(* IEC 61131-3 sources: RVM_Dijital_Ikiz_ModelveOtomasyon_BitirmeProjesi/simulasyon_unity/plc, 14 files *)

(* ---- ST_RVMInput106.st ---- *)
TYPE ST_RVMInput106 :
STRUCT
    uiUnityProtokol : UINT := 106;
    udiUnityOturumu : UDINT := 0;
    udiUnitySayaci : UDINT := 0;
    udiKomutKimligi : UDINT := 0;
    uiOperatorKomutu : UINT := 0;
    xGiris : BOOL := FALSE;
    xTanima : BOOL := FALSE;
    xKiriciGiris : BOOL := FALSE;
    xKirildi : BOOL := FALSE;
    xHazneDolu : BOOL := FALSE;
    xBosaltildi : BOOL := FALSE;
    xKapakAcik : BOOL := FALSE;
    xKapakKapali : BOOL := FALSE;
    xYolBos : BOOL := FALSE;
    xMetalAlgilandi : BOOL := FALSE;
    xSikisma : BOOL := FALSE;
    xAcilStop : BOOL := FALSE;
    xKutuPetDolu : BOOL := FALSE;
    xKutuAluminyumDolu : BOOL := FALSE;
    xKutuCamDolu : BOOL := FALSE;
    rKutleGram : REAL := 0.0;
    rOptikGecirgenlik : REAL := 0.0;
    rBoyMetre : REAL := 0.0;
    rHazneKonumu : REAL := 0.0;
    rGercekBantHizi : REAL := 0.0;
    rGercekKiriciDevri : REAL := 0.0;
    uiBosaltilanKutu : UINT := 0;
    udiUrunKimligi : UDINT := 0;
    uiOperatorParametresi : UINT := 0;
    udiGorulenPlcOturumu : UDINT := 0;
    udiNesneOnayi : UDINT := 0;
    uiNesneSonucu : UINT := 0;
    udiNesneUrunKimligi : UDINT := 0;
    uiPlantVeriKaynagi : UINT := 0;
    xPlantVerisiGecerli : BOOL := FALSE;
    udiGoruntuOnayi : UDINT := 0;
    udiGoruntuUrunu : UDINT := 0;
    udiGoruntuPlcOturumu : UDINT := 0;
    udiGoruntuUnityOturumu : UDINT := 0;
    xGoruntuGecerli : BOOL := FALSE;
    xGoruntuNesneVar : BOOL := FALSE;
    rGoruntuBoy : REAL := 0;
    rGoruntuEn : REAL := 0;
    rGoruntuDoluluk : REAL := 0;
    rGoruntuYasiMs : REAL := 0;
    xOlcumTartiGecerli : BOOL;
    xOlcumProbGecerli : BOOL;
    rOlcumYansima : REAL;
    rOlcumMetal : REAL;
    rOlcumManyetik : REAL;
END_STRUCT
END_TYPE

(* ---- ST_RVMOperator106.st ---- *)
TYPE ST_RVMOperator106 :
STRUCT
    xBaslat : BOOL := FALSE;
    xDurdur : BOOL := FALSE;
    xSifirla : BOOL := FALSE;
    xNesneEkle : BOOL := FALSE;
    xModUygula : BOOL := FALSE;
    xAcilStop : BOOL := FALSE;
    uiSeciliNesne : UINT := 1;
    uiSeciliMod : UINT := 1;
END_STRUCT
END_TYPE

(* ---- ST_RVMOutput106.st ---- *)
TYPE ST_RVMOutput106 :
STRUCT
    uiProtokolSurumu : UINT := 106;
    udiPlcSayaci : UDINT := 0;
    udiUnityOnayOturumu : UDINT := 0;
    udiGirisOnayi : UDINT := 0;
    udiKomutOnayi : UDINT := 0;
    udiIslemKimligi : UDINT := 0;
    uiDurum : UINT := 0;
    uiHataKodu : UINT := 0;
    uiTaninmisMalzeme : UINT := 0;
    uiHedefKutu : UINT := 0;
    xCalismaIzni : BOOL := FALSE;
    xKonveyorIleri : BOOL := FALSE;
    xKonveyorGeri : BOOL := FALSE;
    xKiriciCalis : BOOL := FALSE;
    xHazneHareket : BOOL := FALSE;
    xKapakAc : BOOL := FALSE;
    xTanimaOnayi : BOOL := FALSE;
    rBantHizi : REAL := 0.85;
    rKiriciDevri : REAL := 120.0;
    rHazneHizi : REAL := 1.5;
    rHazneHedefi : REAL := 0.0;
    rKapakAcisi : REAL := 75.0;
    udiPetSayaci : UDINT := 0;
    udiAluminyumSayaci : UDINT := 0;
    udiCamSayaci : UDINT := 0;
    udiReddedilenSayaci : UDINT := 0;
    udiPlcOturumu : UDINT := 0;
    uiKomutDurumu : UINT := 0;
    uiKomutNedeni : UINT := 0;
    udiPlcOperatorKomutKimligi : UDINT := 0;
    uiPlcOperatorKomutu : UINT := 0;
    uiPlcKomutDurumu : UINT := 0;
    uiPlcKomutNedeni : UINT := 0;
    uiSonKomutKaynagi : UINT := 0;
    udiNesneIstegi : UDINT := 0;
    uiNesneProfili : UINT := 0;
    xNesneIstegiEtkin : BOOL := FALSE;
    uiVeriModu : UINT := 1;
    uiDesteklenenModlar : UINT := 2;
    udiCikisBaslangic : UDINT := 0;
    udiCikisBitis : UDINT := 0;
    udiGoruntuIstegi : UDINT := 0;
    uiGoruntuKarari : UINT := 0;
END_STRUCT
END_TYPE

(* ---- GVL_RVMKalici.st ---- *)
{attribute 'qualified_only'}
VAR_GLOBAL PERSISTENT RETAIN
    udiOturum : UDINT;
END_VAR

(* ---- GVL_RVMOperator.st ---- *)
{attribute 'qualified_only'}
VAR_GLOBAL
    xBaslat : BOOL := FALSE;
    xDurdur : BOOL := FALSE;
    xSifirla : BOOL := FALSE;
    xNesneEkle : BOOL := FALSE;
    xModUygula : BOOL := FALSE;
    xAcilStop : BOOL := FALSE;
    uiSeciliNesne : UINT := 1;
    uiSeciliMod : UINT := 1;
END_VAR

(* ---- GVL_RVMUnity.st ---- *)
{attribute 'qualified_only'}
VAR_GLOBAL
    {attribute 'symbol' := 'readwrite'}
    uiUnityProtokol : UINT := 106;
    {attribute 'symbol' := 'readwrite'}
    udiUnityOturumu : UDINT := 0;
    {attribute 'symbol' := 'readwrite'}
    udiUnitySayaci : UDINT := 0;
    {attribute 'symbol' := 'readwrite'}
    udiKomutKimligi : UDINT := 0;
    {attribute 'symbol' := 'readwrite'}
    uiOperatorKomutu : UINT := 0;
    {attribute 'symbol' := 'readwrite'}
    xGiris : BOOL := FALSE;
    {attribute 'symbol' := 'readwrite'}
    xTanima : BOOL := FALSE;
    {attribute 'symbol' := 'readwrite'}
    xKiriciGiris : BOOL := FALSE;
    {attribute 'symbol' := 'readwrite'}
    xKirildi : BOOL := FALSE;
    {attribute 'symbol' := 'readwrite'}
    xHazneDolu : BOOL := FALSE;
    {attribute 'symbol' := 'readwrite'}
    xBosaltildi : BOOL := FALSE;
    {attribute 'symbol' := 'readwrite'}
    xKapakAcik : BOOL := FALSE;
    {attribute 'symbol' := 'readwrite'}
    xKapakKapali : BOOL := FALSE;
    {attribute 'symbol' := 'readwrite'}
    xYolBos : BOOL := FALSE;
    {attribute 'symbol' := 'readwrite'}
    xMetalAlgilandi : BOOL := FALSE;
    {attribute 'symbol' := 'readwrite'}
    xSikisma : BOOL := FALSE;
    {attribute 'symbol' := 'readwrite'}
    xAcilStop : BOOL := FALSE;
    {attribute 'symbol' := 'readwrite'}
    xKutuPetDolu : BOOL := FALSE;
    {attribute 'symbol' := 'readwrite'}
    xKutuAluminyumDolu : BOOL := FALSE;
    {attribute 'symbol' := 'readwrite'}
    xKutuCamDolu : BOOL := FALSE;
    {attribute 'symbol' := 'readwrite'}
    rKutleGram : REAL := 0.0;
    {attribute 'symbol' := 'readwrite'}
    rOptikGecirgenlik : REAL := 0.0;
    {attribute 'symbol' := 'readwrite'}
    rBoyMetre : REAL := 0.0;
    {attribute 'symbol' := 'readwrite'}
    rHazneKonumu : REAL := 0.0;
    {attribute 'symbol' := 'readwrite'}
    rGercekBantHizi : REAL := 0.0;
    {attribute 'symbol' := 'readwrite'}
    rGercekKiriciDevri : REAL := 0.0;
    {attribute 'symbol' := 'readwrite'}
    uiBosaltilanKutu : UINT := 0;
    {attribute 'symbol' := 'readwrite'}
    udiUrunKimligi : UDINT := 0;
    {attribute 'symbol' := 'read'}
    uiProtokolSurumu : UINT := 106;
    {attribute 'symbol' := 'read'}
    udiPlcSayaci : UDINT := 0;
    {attribute 'symbol' := 'read'}
    udiUnityOnayOturumu : UDINT := 0;
    {attribute 'symbol' := 'read'}
    udiGirisOnayi : UDINT := 0;
    {attribute 'symbol' := 'read'}
    udiKomutOnayi : UDINT := 0;
    {attribute 'symbol' := 'read'}
    udiIslemKimligi : UDINT := 0;
    {attribute 'symbol' := 'read'}
    uiDurum : UINT := 0;
    {attribute 'symbol' := 'read'}
    uiHataKodu : UINT := 0;
    {attribute 'symbol' := 'read'}
    uiTaninmisMalzeme : UINT := 0;
    {attribute 'symbol' := 'read'}
    uiHedefKutu : UINT := 0;
    {attribute 'symbol' := 'read'}
    xCalismaIzni : BOOL := FALSE;
    {attribute 'symbol' := 'read'}
    xKonveyorIleri : BOOL := FALSE;
    {attribute 'symbol' := 'read'}
    xKonveyorGeri : BOOL := FALSE;
    {attribute 'symbol' := 'read'}
    xKiriciCalis : BOOL := FALSE;
    {attribute 'symbol' := 'read'}
    xHazneHareket : BOOL := FALSE;
    {attribute 'symbol' := 'read'}
    xKapakAc : BOOL := FALSE;
    {attribute 'symbol' := 'read'}
    xTanimaOnayi : BOOL := FALSE;
    {attribute 'symbol' := 'read'}
    rBantHizi : REAL := 0.85;
    {attribute 'symbol' := 'read'}
    rKiriciDevri : REAL := 120.0;
    {attribute 'symbol' := 'read'}
    rHazneHizi : REAL := 1.5;
    {attribute 'symbol' := 'read'}
    rHazneHedefi : REAL := 0.0;
    {attribute 'symbol' := 'read'}
    rKapakAcisi : REAL := 75.0;
    {attribute 'symbol' := 'read'}
    udiPetSayaci : UDINT := 0;
    {attribute 'symbol' := 'read'}
    udiAluminyumSayaci : UDINT := 0;
    {attribute 'symbol' := 'read'}
    udiCamSayaci : UDINT := 0;
    {attribute 'symbol' := 'read'}
    udiReddedilenSayaci : UDINT := 0;
    {attribute 'symbol' := 'readwrite'}
    udiGirisBaslangic : UDINT := 0;
    {attribute 'symbol' := 'readwrite'}
    udiGirisBitis : UDINT := 0;
    {attribute 'symbol' := 'readwrite'}
    uiOperatorParametresi : UINT := 0;
    {attribute 'symbol' := 'readwrite'}
    udiGorulenPlcOturumu : UDINT := 0;
    {attribute 'symbol' := 'readwrite'}
    udiNesneOnayi : UDINT := 0;
    {attribute 'symbol' := 'readwrite'}
    uiNesneSonucu : UINT := 0;
    {attribute 'symbol' := 'readwrite'}
    udiNesneUrunKimligi : UDINT := 0;
    {attribute 'symbol' := 'readwrite'}
    uiPlantVeriKaynagi : UINT := 0;
    {attribute 'symbol' := 'readwrite'}
    xPlantVerisiGecerli : BOOL := FALSE;
    {attribute 'symbol' := 'read'}
    udiPlcOturumu : UDINT := 0;
    {attribute 'symbol' := 'read'}
    uiKomutDurumu : UINT := 0;
    {attribute 'symbol' := 'read'}
    uiKomutNedeni : UINT := 0;
    {attribute 'symbol' := 'read'}
    udiPlcOperatorKomutKimligi : UDINT := 0;
    {attribute 'symbol' := 'read'}
    uiPlcOperatorKomutu : UINT := 0;
    {attribute 'symbol' := 'read'}
    uiPlcKomutDurumu : UINT := 0;
    {attribute 'symbol' := 'read'}
    uiPlcKomutNedeni : UINT := 0;
    {attribute 'symbol' := 'read'}
    uiSonKomutKaynagi : UINT := 0;
    {attribute 'symbol' := 'read'}
    udiNesneIstegi : UDINT := 0;
    {attribute 'symbol' := 'read'}
    uiNesneProfili : UINT := 0;
    {attribute 'symbol' := 'read'}
    xNesneIstegiEtkin : BOOL := FALSE;
    {attribute 'symbol' := 'read'}
    uiVeriModu : UINT := 1;
    {attribute 'symbol' := 'read'}
    uiDesteklenenModlar : UINT := 2;
    {attribute 'symbol' := 'read'}
    udiCikisBaslangic : UDINT := 0;
    {attribute 'symbol' := 'read'}
    udiCikisBitis : UDINT := 0;
    {attribute 'symbol' := 'readwrite'}
    udiGoruntuOnayi : UDINT := 0;
    {attribute 'symbol' := 'readwrite'}
    udiGoruntuUrunu : UDINT := 0;
    {attribute 'symbol' := 'readwrite'}
    udiGoruntuPlcOturumu : UDINT := 0;
    {attribute 'symbol' := 'readwrite'}
    udiGoruntuUnityOturumu : UDINT := 0;
    {attribute 'symbol' := 'readwrite'}
    xGoruntuGecerli : BOOL := FALSE;
    {attribute 'symbol' := 'readwrite'}
    xGoruntuNesneVar : BOOL := FALSE;
    {attribute 'symbol' := 'readwrite'}
    rGoruntuBoy : REAL := 0;
    {attribute 'symbol' := 'readwrite'}
    rGoruntuEn : REAL := 0;
    {attribute 'symbol' := 'readwrite'}
    rGoruntuDoluluk : REAL := 0;
    {attribute 'symbol' := 'readwrite'}
    rGoruntuYasiMs : REAL := 0;
    {attribute 'symbol' := 'read'}
    udiGoruntuIstegi : UDINT := 0;
    {attribute 'symbol' := 'read'}
    uiGoruntuKarari : UINT := 0;
    {attribute 'symbol' := 'readwrite'}
    xOlcumTartiGecerli : BOOL;
    {attribute 'symbol' := 'readwrite'}
    xOlcumProbGecerli : BOOL;
    {attribute 'symbol' := 'readwrite'}
    rOlcumYansima : REAL;
    {attribute 'symbol' := 'readwrite'}
    rOlcumMetal : REAL;
    {attribute 'symbol' := 'readwrite'}
    rOlcumManyetik : REAL;
END_VAR

(* ---- F_RVMMaterial106_decl.st ---- *)
FUNCTION F_RVMMaterial106 : UINT
VAR_INPUT
    metal : REAL;
    magnetic : REAL;
    grams : REAL;
    transmission : REAL;
    reflection : REAL;
    length : REAL;
    width : REAL;
END_VAR

(* ---- F_RVMPriority106_decl.st ---- *)
FUNCTION F_RVMPriority106 : UINT
VAR_INPUT
    code : UINT;
END_VAR

(* ---- FB_RVMControl106_decl.st ---- *)
FUNCTION_BLOCK FB_RVMControl106
VAR_INPUT
    inp : ST_RVMInput106;
    op : ST_RVMOperator106;
    fresh : BOOL;
    epoch : UDINT;
END_VAR
VAR_OUTPUT
    q : ST_RVMOutput106;
END_VAR
VAR
    a : ST_RVMInput106;
    initialized : BOOL;
    session : UDINT;
    packet : UDINT;
    heartbeat : BOOL;
    synchronized : BOOL;
    sessionChanged : BOOL;
    dataOK : BOOL;
    linked : BOOL;
    home : BOOL;
    emptyHome : BOOL;
    emergency : BOOL;
    stopLevel : BOOL;
    targetFull : BOOL;
    faultNow : UINT;
    previousState : UINT;
    previousButtons : ARRAY[1..5] OF BOOL;
    armed : ARRAY[1..5] OF BOOL;
    buttons : ARRAY[1..5] OF BOOL;
    edges : ARRAY[1..5] OF BOOL;
    newRequest : ARRAY[1..2] OF BOOL;
    cmdId : ARRAY[1..2] OF UDINT;
    cmdCode : ARRAY[1..2] OF UINT;
    cmdParam : ARRAY[1..2] OF UINT;
    cachedStatus : ARRAY[1..2] OF UINT;
    cachedReason : ARRAY[1..2] OF UINT;
    replyId : ARRAY[1..2] OF UDINT;
    replyStatus : ARRAY[1..2] OF UINT;
    replyReason : ARRAY[1..2] OF UINT;
    source : INT;
    chosen : INT;
    other : INT;
    i : INT;
    hmiCode : UINT;
    hmiParam : UINT;
    resultStatus : UINT;
    resultReason : UINT;
    pendingSource : INT;
    pendingId : UDINT;
    insertConfirmed : BOOL;
    confirmedProduct : UDINT;
    lastProduct : UDINT;
    waitLink : TON;
    waitStage : TON;
    waitRecognition : TON;
    waitVision : TON;
    visionMatch : BOOL;
    visionShape : BOOL;
    waitCycle : TON;
    waitInsert : TON;
END_VAR

(* ---- F_RVMMaterial106_body.st ---- *)
// Experimental calibrated rules, not a universal chemical identification.
F_RVMMaterial106 := 0;
IF NOT ((metal>=0) AND (metal<=1) AND (magnetic>=0) AND (magnetic<=0.1)
    AND (grams>=5) AND (grams<=1000) AND (transmission>=0) AND (transmission<=1)
    AND (reflection>=0) AND (reflection<=1) AND (length>=0.10) AND (length<=0.30)
    AND (width>=0.02) AND (width<=0.09)) THEN RETURN; END_IF;
IF metal>=0.5 THEN
    IF (transmission<=0.08) AND (grams>=8) AND (grams<=45) AND (length<=0.20) THEN
        F_RVMMaterial106 := 2;
    END_IF;
ELSIF metal<=0.1 THEN
    IF (grams>=10) AND (grams<=65) AND (transmission>=0.35) THEN F_RVMMaterial106 := 1;
    ELSIF (grams>=100) AND (grams<=800) AND (transmission>=0.15) AND (transmission<=0.85)
        AND (reflection>=0.08) THEN F_RVMMaterial106 := 3;
    END_IF;
END_IF;

(* ---- F_RVMPriority106_body.st ---- *)
CASE code OF
2: F_RVMPriority106 := 1;
3: F_RVMPriority106 := 2;
5: F_RVMPriority106 := 3;
1: F_RVMPriority106 := 4;
4: F_RVMPriority106 := 5;
ELSE F_RVMPriority106 := 99;
END_CASE;

(* ---- FB_RVMControl106_body.st ---- *)
// Single process owner. No actuator command is derived from a UI bit directly.
q.uiProtokolSurumu := 106;
q.udiPlcOturumu := epoch;
q.uiDesteklenenModlar := 2; // Render camera + simulated physical sensors only.
q.uiVeriModu := 1;
q.rBantHizi := 0.85;
q.rKiriciDevri := 120.0;
q.rHazneHizi := 1.5;
q.rKapakAcisi := 75.0;
q.udiPlcSayaci := q.udiPlcSayaci + 1;
heartbeat := FALSE;
sessionChanged := FALSE;
newRequest[1] := FALSE;
newRequest[2] := FALSE;
insertConfirmed := FALSE;
faultNow := 0;
IF NOT initialized THEN
    initialized := TRUE;
    q.uiDurum := 0;
    q.xCalismaIzni := FALSE;
    q.rHazneHedefi := 0.225;
END_IF;
IF epoch = 0 THEN faultNow := 313; END_IF;

// A zero-epoch HELLO is mandatory before this PLC incarnation accepts commands.
// The HELLO'inp command watermark is consumed, never executed.
IF fresh AND (inp.udiUnityOturumu <> 0) AND (inp.udiUnitySayaci <> 0) THEN
    IF (inp.udiGorulenPlcOturumu = 0) AND ((session <> inp.udiUnityOturumu) OR NOT synchronized) THEN
        a := inp;
        sessionChanged := session <> inp.udiUnityOturumu;
        session := inp.udiUnityOturumu;
        lastProduct := 0;
        packet := inp.udiUnitySayaci;
        synchronized := TRUE;
        cmdId[1] := inp.udiKomutKimligi;
        cmdCode[1] := inp.uiOperatorKomutu;
        cmdParam[1] := inp.uiOperatorParametresi;
        cachedStatus[1] := 5;
        cachedReason[1] := 10;
        replyId[1] := cmdId[1];
        replyStatus[1] := 5;
        replyReason[1] := 10;
        q.xCalismaIzni := FALSE;
        IF q.uiHataKodu = 0 THEN q.uiDurum := 0; END_IF;
    ELSIF synchronized AND (session = inp.udiUnityOturumu)
        AND (inp.udiGorulenPlcOturumu = epoch) AND (inp.udiUnitySayaci > packet) THEN
        packet := inp.udiUnitySayaci;
        a := inp;
        heartbeat := TRUE;
        IF inp.udiKomutKimligi > cmdId[1] THEN
            cmdId[1] := inp.udiKomutKimligi;
            cmdCode[1] := inp.uiOperatorKomutu;
            cmdParam[1] := inp.uiOperatorParametresi;
            newRequest[1] := TRUE;
        ELSIF (inp.udiKomutKimligi <> cmdId[1]) OR (inp.uiOperatorKomutu <> cmdCode[1])
            OR (inp.uiOperatorParametresi <> cmdParam[1]) THEN
            replyId[1] := inp.udiKomutKimligi;
            replyStatus[1] := 3;
            replyReason[1] := 13;
        ELSE
            replyId[1] := cmdId[1];
            replyStatus[1] := cachedStatus[1];
            replyReason[1] := cachedReason[1];
        END_IF;
    END_IF;
END_IF;
q.udiUnityOnayOturumu := session;
waitLink(IN := NOT heartbeat, PT := T#750MS);
linked := synchronized AND (session = a.udiUnityOturumu) AND (a.udiGorulenPlcOturumu = epoch)
    AND (epoch <> 0) AND NOT waitLink.Q AND (a.uiUnityProtokol = 106);
home := ABS(a.rHazneKonumu - 0.225) < 0.008;
emptyHome := a.xYolBos AND NOT a.xGiris AND a.xKapakKapali AND NOT a.xKapakAcik AND home;
emergency := op.xAcilStop OR a.xAcilStop;
// Comparisons reject NaN as well as out-of-range values. No invalid data fallback.
dataOK := a.xPlantVerisiGecerli AND (a.uiPlantVeriKaynagi = 1)
    AND (a.rHazneKonumu >= -0.770001) AND (a.rHazneKonumu <= 0.310001)
    AND (a.rKutleGram >= 0.0) AND (a.rKutleGram <= 10000.0)
    AND (a.rBoyMetre >= 0.0) AND (a.rBoyMetre <= 2.000001)
    AND (a.rOptikGecirgenlik >= 0.0) AND (a.rOptikGecirgenlik <= 1.000001)
    AND (a.rGercekBantHizi >= -1.200001) AND (a.rGercekBantHizi <= 1.200001)
    AND (a.rGercekKiriciDevri >= 0.0) AND (a.rGercekKiriciDevri <= 180.0001)
    AND NOT (a.xKapakAcik AND a.xKapakKapali)
    AND NOT (a.xYolBos AND a.xGiris) AND (a.uiBosaltilanKutu <= 3);

// HMI: arm only after FALSE has been observed; held or startup TRUE cannot repeat.
buttons[1] := op.xBaslat; buttons[2] := op.xDurdur; buttons[3] := op.xSifirla;
buttons[4] := op.xNesneEkle; buttons[5] := op.xModUygula;
FOR i := 1 TO 5 DO
    IF NOT buttons[i] THEN armed[i] := TRUE; END_IF;
    edges[i] := armed[i] AND buttons[i] AND NOT previousButtons[i];
    previousButtons[i] := buttons[i];
END_FOR;
hmiCode := 0; hmiParam := 0;
IF edges[2] THEN hmiCode := 2;
ELSIF edges[3] THEN hmiCode := 3;
ELSIF edges[5] THEN hmiCode := 5; hmiParam := op.uiSeciliMod;
ELSIF edges[1] THEN hmiCode := 1;
ELSIF edges[4] THEN hmiCode := 4; hmiParam := op.uiSeciliNesne;
END_IF;
IF hmiCode <> 0 THEN
    IF cmdId[2] = UDINT#4294967295 THEN faultNow := 313;
    ELSE
        cmdId[2] := cmdId[2] + 1;
        cmdCode[2] := hmiCode; cmdParam[2] := hmiParam;
        newRequest[2] := TRUE;
    END_IF;
END_IF;
stopLevel := op.xDurdur OR (newRequest[1] AND (cmdCode[1] = 2));

// Fault priority is stable; reconnecting Unity never clears a latched fault.
IF q.xCalismaIzni THEN
    IF emergency THEN faultNow := 303;
    // Unity also raises its local motion interlock on an identity mismatch.
    // Preserve the specific cause while the session is valid, before generic jam/data flags.
    ELSIF linked AND (q.uiDurum >= 20) AND (q.uiDurum <= 100) AND (a.udiUrunKimligi <> q.udiIslemKimligi) THEN faultNow := 305;
    ELSIF a.xSikisma THEN faultNow := 304;
    ELSIF a.uiUnityProtokol <> 106 THEN faultNow := 302;
    ELSIF NOT linked THEN faultNow := 301;
    ELSIF NOT dataOK THEN faultNow := 310;
    END_IF;
END_IF;
waitStage(IN := (q.uiDurum = previousState) AND (q.uiDurum >= 20) AND (q.uiDurum <= 100), PT := T#8S);
previousState := q.uiDurum;
waitRecognition(IN := q.uiDurum = 30, PT := T#200MS);
waitVision(IN := q.uiDurum = 30, PT := T#4S);
visionMatch := (a.udiGoruntuOnayi = q.udiGoruntuIstegi) AND (q.udiGoruntuIstegi <> 0)
    AND (a.udiGoruntuUrunu = q.udiIslemKimligi) AND (a.udiGoruntuPlcOturumu = epoch)
    AND (a.udiGoruntuUnityOturumu = session);
visionShape := a.xGoruntuNesneVar AND (a.rGoruntuBoy >= 0.10) AND (a.rGoruntuBoy <= 0.30)
    AND (a.rGoruntuEn >= 0.02) AND (a.rGoruntuEn <= 0.09)
    AND (a.rGoruntuBoy >= 1.5*a.rGoruntuEn) AND (a.rGoruntuBoy <= 7.0*a.rGoruntuEn)
    AND (a.rGoruntuDoluluk >= 0.35) AND (a.rGoruntuDoluluk <= 1.0);
waitCycle(IN := (q.uiDurum >= 20) AND (q.uiDurum <= 90), PT := T#5600MS);
waitInsert(IN := q.xNesneIstegiEtkin, PT := T#2S);
IF waitStage.Q AND (faultNow = 0) THEN faultNow := 306; END_IF;
IF faultNow <> 0 AND q.uiHataKodu = 0 THEN q.uiHataKodu := faultNow; END_IF;
IF stopLevel OR emergency OR sessionChanged OR (q.uiHataKodu <> 0) THEN
    q.xCalismaIzni := FALSE;
    IF q.uiHataKodu = 0 THEN q.uiDurum := 0; ELSE q.uiDurum := 900; END_IF;
    IF q.xNesneIstegiEtkin THEN
        cachedStatus[pendingSource] := 5; cachedReason[pendingSource] := 1;
        IF replyId[pendingSource] = pendingId THEN
            replyStatus[pendingSource] := 5; replyReason[pendingSource] := 1;
        END_IF;
    END_IF;
    q.xNesneIstegiEtkin := FALSE;
END_IF;

// Arbitration is deterministic. No deferred queue can start work after a stop.
chosen := 0;
IF newRequest[2] THEN chosen := 2; END_IF;
IF newRequest[1] THEN
    IF chosen = 0 THEN chosen := 1;
    ELSIF F_RVMPriority106(cmdCode[1]) < F_RVMPriority106(cmdCode[2]) THEN chosen := 1;
    END_IF;
END_IF;
FOR source := 1 TO 2 DO
    IF newRequest[source] THEN
        resultStatus := 3; resultReason := 0;
        replyId[source] := cmdId[source];
        IF (source <> chosen) AND NOT (cmdCode[source] = 2) THEN
            IF stopLevel THEN resultReason := 1; ELSE resultReason := 9; END_IF;
        ELSIF cmdCode[source] = 2 THEN
            q.xCalismaIzni := FALSE;
            IF q.uiHataKodu = 0 THEN q.uiDurum := 0; ELSE q.uiDurum := 900; END_IF;
            resultStatus := 2;
        ELSIF (cmdCode[source] = 0) OR (cmdCode[source] > 5)
            OR ((cmdCode[source] <= 3) AND (cmdParam[source] <> 0))
            OR ((cmdCode[source] = 4) AND (cmdParam[source] > 3))
            OR ((cmdCode[source] = 5) AND (cmdParam[source] > 2)) THEN resultReason := 7;
        ELSIF stopLevel THEN resultReason := 1;
        ELSIF emergency OR a.xSikisma THEN resultReason := 5;
        ELSIF NOT linked OR NOT dataOK THEN resultReason := 2;
        ELSIF q.xNesneIstegiEtkin THEN resultReason := 6;
        ELSE
            CASE cmdCode[source] OF
            1:
                IF q.uiHataKodu <> 0 THEN resultReason := 5;
                ELSIF q.uiDurum <> 0 THEN resultReason := 3;
                ELSIF NOT emptyHome THEN resultReason := 4;
                ELSE q.xCalismaIzni := TRUE; q.uiDurum := 10; resultStatus := 2;
                END_IF;
            3:
                IF q.xCalismaIzni OR ((q.uiDurum <> 0) AND (q.uiDurum <> 900)) THEN resultReason := 3;
                ELSIF NOT emptyHome THEN resultReason := 4;
                ELSIF epoch = 0 THEN resultReason := 10;
                ELSE q.uiHataKodu := 0; q.uiDurum := 0; q.xCalismaIzni := FALSE; resultStatus := 2;
                END_IF;
            4:
                IF q.uiHataKodu <> 0 THEN resultReason := 5;
                ELSIF (q.uiDurum <> 10) OR NOT q.xCalismaIzni THEN resultReason := 3;
                ELSIF NOT emptyHome THEN resultReason := 4;
                ELSIF q.udiNesneIstegi = UDINT#4294967295 THEN resultReason := 10;
                ELSE
                    q.udiNesneIstegi := q.udiNesneIstegi + 1;
                    q.uiNesneProfili := cmdParam[source];
                    q.xNesneIstegiEtkin := TRUE;
                    pendingSource := source; pendingId := cmdId[source];
                    resultStatus := 1;
                END_IF;
            5:
                IF cmdParam[source] <> 1 THEN resultReason := 8;
                ELSIF (q.uiDurum <> 0) OR q.xCalismaIzni THEN resultReason := 3;
                ELSIF NOT emptyHome THEN resultReason := 4;
                ELSE q.uiVeriModu := 1; resultStatus := 2;
                END_IF;
            END_CASE;
        END_IF;
        cachedStatus[source] := resultStatus; cachedReason[source] := resultReason;
        replyStatus[source] := resultStatus; replyReason[source] := resultReason;
        IF source = chosen THEN q.uiSonKomutKaynagi := INT_TO_UINT(source); END_IF;
    END_IF;
END_FOR;

// Product admission is tied to the PLC-issued request, not just a presence bit.
IF q.xNesneIstegiEtkin THEN
    resultStatus := 1; resultReason := 0;
    IF waitInsert.Q THEN
        resultStatus := 4; resultReason := 11;
        q.uiHataKodu := 312; // A delayed physical creation must require explicit recovery.
    ELSIF heartbeat AND (a.udiNesneOnayi = q.udiNesneIstegi) THEN
        IF a.uiNesneSonucu = 2 THEN resultStatus := 3; resultReason := 12;
        ELSIF a.uiNesneSonucu = 1 THEN
            IF (a.udiNesneUrunKimligi <> 0) AND (a.udiNesneUrunKimligi = a.udiUrunKimligi)
                AND (a.udiUrunKimligi > lastProduct) AND a.xGiris AND NOT a.xYolBos THEN
                confirmedProduct := a.udiUrunKimligi;
                lastProduct := a.udiUrunKimligi;
                insertConfirmed := TRUE;
                resultStatus := 2;
            ELSE resultStatus := 3; resultReason := 12; q.uiHataKodu := 312;
            END_IF;
        END_IF;
    END_IF;
    IF resultStatus <> 1 THEN
        q.xNesneIstegiEtkin := FALSE;
        IF cmdId[pendingSource] = pendingId THEN
            cachedStatus[pendingSource] := resultStatus; cachedReason[pendingSource] := resultReason;
        END_IF;
        IF replyId[pendingSource] = pendingId THEN
            replyStatus[pendingSource] := resultStatus; replyReason[pendingSource] := resultReason;
        END_IF;
    END_IF;
END_IF;

targetFull := ((q.uiHedefKutu = 1) AND a.xKutuPetDolu)
    OR ((q.uiHedefKutu = 2) AND a.xKutuAluminyumDolu)
    OR ((q.uiHedefKutu = 3) AND a.xKutuCamDolu);
IF q.xCalismaIzni AND (q.uiDurum >= 40) AND (q.uiDurum <= 70) AND targetFull THEN q.uiHataKodu := 308; END_IF;
IF q.uiHataKodu = 0 AND q.xCalismaIzni THEN
    CASE q.uiDurum OF
    10:
        q.xTanimaOnayi := FALSE; q.uiTaninmisMalzeme := 0; q.uiHedefKutu := 0;
        IF insertConfirmed THEN q.udiIslemKimligi := confirmedProduct; q.uiDurum := 20;
        ELSIF NOT a.xYolBos AND NOT q.xNesneIstegiEtkin THEN q.uiHataKodu := 312;
        END_IF;
    20:
        IF a.xTanima THEN
            IF q.udiGoruntuIstegi = UDINT#4294967295 THEN q.uiHataKodu := 313;
            ELSE q.udiGoruntuIstegi := q.udiGoruntuIstegi+1; q.uiGoruntuKarari := 0; q.uiDurum := 30;
            END_IF;
        END_IF;
    30:
        IF NOT a.xTanima THEN q.uiHataKodu := 307;
        ELSIF waitVision.Q THEN
            q.uiGoruntuKarari := 5; q.uiTaninmisMalzeme := 0; q.uiHedefKutu := 0; q.uiDurum := 100;
        ELSIF waitRecognition.Q AND visionMatch THEN
            q.uiTaninmisMalzeme := 0;
            IF NOT ((a.rGoruntuYasiMs >= 0.0) AND (a.rGoruntuYasiMs <= 2000.0)) THEN q.uiGoruntuKarari := 4;
            ELSIF NOT a.xGoruntuGecerli OR NOT a.xOlcumTartiGecerli OR NOT a.xOlcumProbGecerli THEN q.uiGoruntuKarari := 3;
            ELSIF NOT visionShape THEN q.uiGoruntuKarari := 2;
            ELSE
                q.uiTaninmisMalzeme := F_RVMMaterial106(a.rOlcumMetal, a.rOlcumManyetik, a.rKutleGram, a.rOptikGecirgenlik, a.rOlcumYansima, a.rGoruntuBoy, a.rGoruntuEn);
                IF q.uiTaninmisMalzeme = 0 THEN q.uiGoruntuKarari := 2; ELSE q.uiGoruntuKarari := 1; END_IF;
            END_IF;
            q.uiHedefKutu := q.uiTaninmisMalzeme;
            CASE q.uiHedefKutu OF
            1: q.rHazneHedefi := -0.23;
            2: q.rHazneHedefi := -0.77;
            3: q.rHazneHedefi := 0.31;
            END_CASE;
            IF q.uiHedefKutu = 0 THEN q.uiDurum := 100;
            ELSIF ((q.uiHedefKutu=1) AND a.xKutuPetDolu) OR ((q.uiHedefKutu=2) AND a.xKutuAluminyumDolu)
                OR ((q.uiHedefKutu=3) AND a.xKutuCamDolu) THEN q.uiHataKodu := 308;
            ELSE q.xTanimaOnayi := TRUE; q.uiDurum := 40;
            END_IF;
        END_IF;
    40:
        IF NOT a.xKapakKapali THEN q.uiHataKodu := 310;
        ELSIF a.xKiriciGiris THEN q.uiDurum := 50; END_IF;
    50:
        IF a.xKirildi AND a.xHazneDolu AND a.xKapakKapali THEN q.uiDurum := 60; END_IF;
    60:
        IF NOT a.xKapakKapali OR NOT a.xHazneDolu THEN q.uiHataKodu := 310;
        ELSIF ABS(a.rHazneKonumu-q.rHazneHedefi)<0.008 THEN q.uiDurum := 70; END_IF;
    70:
        IF ABS(a.rHazneKonumu-q.rHazneHedefi)>=0.008 THEN q.uiHataKodu := 310;
        ELSIF a.xBosaltildi AND a.xKapakAcik AND NOT a.xHazneDolu AND a.xYolBos THEN
            IF a.uiBosaltilanKutu <> q.uiHedefKutu THEN q.uiHataKodu := 309;
            ELSE q.uiDurum := 80; END_IF;
        END_IF;
    80:
        IF a.xKapakKapali AND NOT a.xKapakAcik AND a.xYolBos AND NOT a.xHazneDolu THEN
            CASE q.uiHedefKutu OF
            1: q.udiPetSayaci := q.udiPetSayaci + 1;
            2: q.udiAluminyumSayaci := q.udiAluminyumSayaci + 1;
            3: q.udiCamSayaci := q.udiCamSayaci + 1;
            END_CASE;
            q.uiDurum := 90;
        END_IF;
    90:
        q.rHazneHedefi := 0.225;
        IF NOT a.xKapakKapali THEN q.uiHataKodu := 310;
        ELSIF home AND a.xYolBos AND waitCycle.Q THEN q.uiDurum := 10; END_IF;
    100:
        IF a.xYolBos THEN q.udiReddedilenSayaci := q.udiReddedilenSayaci+1; q.uiDurum := 10; END_IF;
    END_CASE;
END_IF;

// Apply fault dominance AFTER state processing, in this same scan.
IF q.uiHataKodu <> 0 THEN q.uiDurum := 900; q.xCalismaIzni := FALSE; q.xNesneIstegiEtkin := FALSE; END_IF;
q.xKonveyorIleri := FALSE; q.xKonveyorGeri := FALSE; q.xKiriciCalis := FALSE;
q.xHazneHareket := FALSE; q.xKapakAc := FALSE;
IF q.xCalismaIzni AND linked AND dataOK AND NOT emergency AND NOT a.xSikisma AND NOT stopLevel THEN
    q.xKonveyorIleri := (q.uiDurum=20) OR (q.uiDurum=40);
    q.xKonveyorGeri := q.uiDurum=100;
    q.xKiriciCalis := ((q.uiDurum=40) OR (q.uiDurum=50)) AND q.xTanimaOnayi;
    q.xHazneHareket := ((q.uiDurum=60) OR (q.uiDurum=90)) AND a.xKapakKapali;
    q.xKapakAc := (q.uiDurum=70) AND (ABS(a.rHazneKonumu-q.rHazneHedefi)<0.008);
END_IF;
IF NOT q.xCalismaIzni THEN q.xTanimaOnayi := FALSE; END_IF;
q.udiKomutOnayi := replyId[1]; q.uiKomutDurumu := replyStatus[1]; q.uiKomutNedeni := replyReason[1];
q.udiPlcOperatorKomutKimligi := replyId[2]; q.uiPlcOperatorKomutu := cmdCode[2];
q.uiPlcKomutDurumu := replyStatus[2]; q.uiPlcKomutNedeni := replyReason[2];

(* ---- PRG_UnityRVM_body.st ---- *)
IF NOT initialized THEN
    initialized := TRUE;
    IF GVL_RVMKalici.udiOturum < UDINT#4294967295 THEN
        GVL_RVMKalici.udiOturum := GVL_RVMKalici.udiOturum + 1;
        epoch := GVL_RVMKalici.udiOturum;
    END_IF;
END_IF;
fresh := FALSE;
beginMarker := GVL_RVMUnity.udiGirisBaslangic;
IF (beginMarker <> 0) AND (beginMarker = GVL_RVMUnity.udiGirisBitis) AND (beginMarker <> lastMarker) THEN
candidate.uiUnityProtokol := GVL_RVMUnity.uiUnityProtokol;
candidate.udiUnityOturumu := GVL_RVMUnity.udiUnityOturumu;
candidate.udiUnitySayaci := GVL_RVMUnity.udiUnitySayaci;
candidate.udiKomutKimligi := GVL_RVMUnity.udiKomutKimligi;
candidate.uiOperatorKomutu := GVL_RVMUnity.uiOperatorKomutu;
candidate.xGiris := GVL_RVMUnity.xGiris;
candidate.xTanima := GVL_RVMUnity.xTanima;
candidate.xKiriciGiris := GVL_RVMUnity.xKiriciGiris;
candidate.xKirildi := GVL_RVMUnity.xKirildi;
candidate.xHazneDolu := GVL_RVMUnity.xHazneDolu;
candidate.xBosaltildi := GVL_RVMUnity.xBosaltildi;
candidate.xKapakAcik := GVL_RVMUnity.xKapakAcik;
candidate.xKapakKapali := GVL_RVMUnity.xKapakKapali;
candidate.xYolBos := GVL_RVMUnity.xYolBos;
candidate.xMetalAlgilandi := GVL_RVMUnity.xMetalAlgilandi;
candidate.xSikisma := GVL_RVMUnity.xSikisma;
candidate.xAcilStop := GVL_RVMUnity.xAcilStop;
candidate.xKutuPetDolu := GVL_RVMUnity.xKutuPetDolu;
candidate.xKutuAluminyumDolu := GVL_RVMUnity.xKutuAluminyumDolu;
candidate.xKutuCamDolu := GVL_RVMUnity.xKutuCamDolu;
candidate.rKutleGram := GVL_RVMUnity.rKutleGram;
candidate.rOptikGecirgenlik := GVL_RVMUnity.rOptikGecirgenlik;
candidate.rBoyMetre := GVL_RVMUnity.rBoyMetre;
candidate.rHazneKonumu := GVL_RVMUnity.rHazneKonumu;
candidate.rGercekBantHizi := GVL_RVMUnity.rGercekBantHizi;
candidate.rGercekKiriciDevri := GVL_RVMUnity.rGercekKiriciDevri;
candidate.uiBosaltilanKutu := GVL_RVMUnity.uiBosaltilanKutu;
candidate.udiUrunKimligi := GVL_RVMUnity.udiUrunKimligi;
candidate.uiOperatorParametresi := GVL_RVMUnity.uiOperatorParametresi;
candidate.udiGorulenPlcOturumu := GVL_RVMUnity.udiGorulenPlcOturumu;
candidate.udiNesneOnayi := GVL_RVMUnity.udiNesneOnayi;
candidate.uiNesneSonucu := GVL_RVMUnity.uiNesneSonucu;
candidate.udiNesneUrunKimligi := GVL_RVMUnity.udiNesneUrunKimligi;
candidate.uiPlantVeriKaynagi := GVL_RVMUnity.uiPlantVeriKaynagi;
candidate.xPlantVerisiGecerli := GVL_RVMUnity.xPlantVerisiGecerli;
candidate.udiGoruntuOnayi := GVL_RVMUnity.udiGoruntuOnayi;
candidate.udiGoruntuUrunu := GVL_RVMUnity.udiGoruntuUrunu;
candidate.udiGoruntuPlcOturumu := GVL_RVMUnity.udiGoruntuPlcOturumu;
candidate.udiGoruntuUnityOturumu := GVL_RVMUnity.udiGoruntuUnityOturumu;
candidate.xGoruntuGecerli := GVL_RVMUnity.xGoruntuGecerli;
candidate.xGoruntuNesneVar := GVL_RVMUnity.xGoruntuNesneVar;
candidate.rGoruntuBoy := GVL_RVMUnity.rGoruntuBoy;
candidate.rGoruntuEn := GVL_RVMUnity.rGoruntuEn;
candidate.rGoruntuDoluluk := GVL_RVMUnity.rGoruntuDoluluk;
candidate.rGoruntuYasiMs := GVL_RVMUnity.rGoruntuYasiMs;
candidate.xOlcumTartiGecerli := GVL_RVMUnity.xOlcumTartiGecerli;
candidate.xOlcumProbGecerli := GVL_RVMUnity.xOlcumProbGecerli;
candidate.rOlcumYansima := GVL_RVMUnity.rOlcumYansima;
candidate.rOlcumMetal := GVL_RVMUnity.rOlcumMetal;
candidate.rOlcumManyetik := GVL_RVMUnity.rOlcumManyetik;
    fresh := (beginMarker = GVL_RVMUnity.udiGirisBitis) AND (beginMarker = GVL_RVMUnity.udiGirisBaslangic);
    IF fresh THEN snapshot := candidate; lastMarker := beginMarker; END_IF;
END_IF;
op.xBaslat := GVL_RVMOperator.xBaslat;
op.xDurdur := GVL_RVMOperator.xDurdur;
op.xSifirla := GVL_RVMOperator.xSifirla;
op.xNesneEkle := GVL_RVMOperator.xNesneEkle;
op.xModUygula := GVL_RVMOperator.xModUygula;
op.xAcilStop := GVL_RVMOperator.xAcilStop;
op.uiSeciliNesne := GVL_RVMOperator.uiSeciliNesne;
op.uiSeciliMod := GVL_RVMOperator.uiSeciliMod;
control(inp := snapshot, op := op, fresh := fresh, epoch := epoch);
IF outputMarker = UDINT#4294967295 THEN outputMarker := 1; ELSE outputMarker := outputMarker+1; END_IF;
GVL_RVMUnity.udiCikisBaslangic := outputMarker;
GVL_RVMUnity.uiProtokolSurumu := control.q.uiProtokolSurumu;
GVL_RVMUnity.udiPlcSayaci := control.q.udiPlcSayaci;
GVL_RVMUnity.udiUnityOnayOturumu := control.q.udiUnityOnayOturumu;
GVL_RVMUnity.udiGirisOnayi := control.q.udiGirisOnayi;
GVL_RVMUnity.udiKomutOnayi := control.q.udiKomutOnayi;
GVL_RVMUnity.udiIslemKimligi := control.q.udiIslemKimligi;
GVL_RVMUnity.uiDurum := control.q.uiDurum;
GVL_RVMUnity.uiHataKodu := control.q.uiHataKodu;
GVL_RVMUnity.uiTaninmisMalzeme := control.q.uiTaninmisMalzeme;
GVL_RVMUnity.uiHedefKutu := control.q.uiHedefKutu;
GVL_RVMUnity.xCalismaIzni := control.q.xCalismaIzni;
GVL_RVMUnity.xKonveyorIleri := control.q.xKonveyorIleri;
GVL_RVMUnity.xKonveyorGeri := control.q.xKonveyorGeri;
GVL_RVMUnity.xKiriciCalis := control.q.xKiriciCalis;
GVL_RVMUnity.xHazneHareket := control.q.xHazneHareket;
GVL_RVMUnity.xKapakAc := control.q.xKapakAc;
GVL_RVMUnity.xTanimaOnayi := control.q.xTanimaOnayi;
GVL_RVMUnity.rBantHizi := control.q.rBantHizi;
GVL_RVMUnity.rKiriciDevri := control.q.rKiriciDevri;
GVL_RVMUnity.rHazneHizi := control.q.rHazneHizi;
GVL_RVMUnity.rHazneHedefi := control.q.rHazneHedefi;
GVL_RVMUnity.rKapakAcisi := control.q.rKapakAcisi;
GVL_RVMUnity.udiPetSayaci := control.q.udiPetSayaci;
GVL_RVMUnity.udiAluminyumSayaci := control.q.udiAluminyumSayaci;
GVL_RVMUnity.udiCamSayaci := control.q.udiCamSayaci;
GVL_RVMUnity.udiReddedilenSayaci := control.q.udiReddedilenSayaci;
GVL_RVMUnity.udiPlcOturumu := control.q.udiPlcOturumu;
GVL_RVMUnity.uiKomutDurumu := control.q.uiKomutDurumu;
GVL_RVMUnity.uiKomutNedeni := control.q.uiKomutNedeni;
GVL_RVMUnity.udiPlcOperatorKomutKimligi := control.q.udiPlcOperatorKomutKimligi;
GVL_RVMUnity.uiPlcOperatorKomutu := control.q.uiPlcOperatorKomutu;
GVL_RVMUnity.uiPlcKomutDurumu := control.q.uiPlcKomutDurumu;
GVL_RVMUnity.uiPlcKomutNedeni := control.q.uiPlcKomutNedeni;
GVL_RVMUnity.uiSonKomutKaynagi := control.q.uiSonKomutKaynagi;
GVL_RVMUnity.udiNesneIstegi := control.q.udiNesneIstegi;
GVL_RVMUnity.uiNesneProfili := control.q.uiNesneProfili;
GVL_RVMUnity.xNesneIstegiEtkin := control.q.xNesneIstegiEtkin;
GVL_RVMUnity.uiVeriModu := control.q.uiVeriModu;
GVL_RVMUnity.uiDesteklenenModlar := control.q.uiDesteklenenModlar;
GVL_RVMUnity.udiGoruntuIstegi := control.q.udiGoruntuIstegi;
GVL_RVMUnity.uiGoruntuKarari := control.q.uiGoruntuKarari;
GVL_RVMUnity.udiGirisOnayi := lastMarker;
GVL_RVMUnity.udiCikisBitis := outputMarker;

(* ---- PRG_UnityRVM_decl.st ---- *)
PROGRAM PRG_UnityRVM
VAR
    control : FB_RVMControl106;
    candidate : ST_RVMInput106;
    snapshot : ST_RVMInput106;
    op : ST_RVMOperator106;
    initialized : BOOL;
    epoch : UDINT;
    beginMarker : UDINT;
    lastMarker : UDINT;
    outputMarker : UDINT;
    fresh : BOOL;
END_VAR
